(* IEC 61131-3 sources: botanik2/src/libbotanik/plc/functions, 5 files *)

(* ---- health.st ---- *)
(* What a program says about its own answer
   ------------------------------------------------------------------------ *)

(* The codes are Plc::Health's, in its order: matiec numbers an enumeration
   0,1,2... in declaration order, and the two sides have to agree because the
   value IS the program's health row. matiec rejects explicit values here, so
   the order is the contract.

   Only a program that OPTS IN (`health` in programs.csv) has a row to write,
   and one that opts in owes a write to it on every path - which the generator
   checks off matiec's own write list, the same way it checks a quality.

   Every output is written on every scan, so this is never about whether a row
   moved. It is what the number MEANS. *)

TYPE
  HEALTH : (HEALTHY, DEGRADED, FAULTED);
END_TYPE

FUNCTION WORST_HEALTH : HEALTH
(* How a program that leans on another's answer inherits it: the weaker of the
   two. Spelled as comparisons rather than as a maximum, because the ordering
   of an enumerated type is not something to lean on. *)
VAR_INPUT
  A : HEALTH;
  B : HEALTH;
END_VAR
  IF A = FAULTED OR B = FAULTED THEN WORST_HEALTH := FAULTED;
  ELSIF A = DEGRADED OR B = DEGRADED THEN WORST_HEALTH := DEGRADED;
  ELSE WORST_HEALTH := HEALTHY; END_IF;
END_FUNCTION

FUNCTION VERDICT : HEALTH
(* The common shape, said once: whether the law could answer at all, and
   whether it trusted what it answered on.

   ANSWERED is asked first and separately because the two are not degrees of
   one thing: a law with no evidence at all writes its safe state, which is a
   different fact from a law that chose a fallback and stands behind it. *)
VAR_INPUT
  ANSWERED : BOOL;
  TRUSTED  : BOOL;
END_VAR
  IF NOT ANSWERED THEN VERDICT := FAULTED;
  ELSIF NOT TRUSTED THEN VERDICT := DEGRADED;
  ELSE VERDICT := HEALTHY; END_IF;
END_FUNCTION

(* ---- quality.st ---- *)
(* What a reading is worth, and the two ways a law asks
   ------------------------------------------------------------------------ *)

(* The codes are Vars::Quality's, in its order: matiec numbers an enumeration
   0,1,2... in declaration order, and the two sides have to agree because the
   value IS the companion row's. matiec rejects explicit values here, so the
   order is the contract.

   Three, and each is a DECISION a reader makes differently: nothing behind the
   row, something measured, or a number the law stands behind though nothing
   measured it. The reasons a reading went bad - stale, out of band, refused -
   are diagnoses rather than decisions, and each has a home of its own: the
   stamp's age, the band beside the value, and one log line from the master. *)

TYPE
  QUALITY : (Q_NONE, Q_GOOD, Q_HELD);
END_TYPE

FUNCTION GOOD : BOOL
(* Whether something MEASURED it. What a law gating on seeing the plant asks. *)
VAR_INPUT
  Q : QUALITY;
END_VAR
  GOOD := Q = Q_GOOD;
END_FUNCTION

FUNCTION USABLE : BOOL
(* Whether there is a NUMBER behind it worth computing on. Wider than GOOD by
   exactly Q_HELD, which is a law's own fallback. *)
VAR_INPUT
  Q : QUALITY;
END_VAR
  USABLE := Q <> Q_NONE;
END_FUNCTION

FUNCTION WORST_OF : QUALITY
(* How a derived row inherits its inputs': the weaker of the two. Spelled as
   comparisons rather than as a minimum, because the ordering of an enumerated
   type is not something to lean on. *)
VAR_INPUT
  A : QUALITY;
  B : QUALITY;
END_VAR
  IF A = Q_NONE OR B = Q_NONE THEN WORST_OF := Q_NONE;
  ELSIF A = Q_HELD OR B = Q_HELD THEN WORST_OF := Q_HELD;
  ELSE WORST_OF := Q_GOOD; END_IF;
END_FUNCTION

FUNCTION QUAL : QUALITY
(* The quality of a row a law publishes with no input verdict to inherit:
   measured this beat, HOLDING something it measured once, or nothing it has
   ever seen.

   SEEDED is asked separately and always, because the middle case is the one
   that gets skipped: a block whose output holds its last reading and reports
   only OK publishes Q_NONE for a row that has real evidence in it, and
   Ref::get() then hands every reader the declared value instead. Pass FALSE
   where the law genuinely holds nothing - a verdict recomputed each scan - and
   let that be a claim somebody made rather than a default. *)
VAR_INPUT
  OK     : BOOL;
  SEEDED : BOOL;
END_VAR
  IF OK THEN QUAL := Q_GOOD;
  ELSIF SEEDED THEN QUAL := Q_HELD;
  ELSE QUAL := Q_NONE; END_IF;
END_FUNCTION

(* ---- math.st ---- *)
(* The demand ladders, and the votes a redundant chain reduces with
   ------------------------------------------------------------------------ *)

(* Written once so three subsystems cannot disagree about what "half demand"
   means. Stateless, so FUNCTIONs rather than blocks. *)

FUNCTION LADDER : REAL
(* V mapped onto 0..1 across [LO, HI] and clamped. A degenerate or inverted
   span reads as fully on at or above HI, so a mis-set pair fails toward
   ACTING rather than toward doing nothing. *)
VAR_INPUT
  V  : REAL;
  LO : REAL;
  HI : REAL;
END_VAR
  IF HI <= LO THEN
    IF V >= HI THEN LADDER := 1.0; ELSE LADDER := 0.0; END_IF;
  ELSE
    LADDER := LIMIT(0.0, (V - LO) / (HI - LO), 1.0);
  END_IF;
END_FUNCTION

FUNCTION SIGNED_LADDER : REAL
(* The same either side of zero, with a dead band between. Reads 0 inside
   [NEG_START, POS_START], falls to -1 by NEG_FULL and rises to +1 by
   POS_FULL. One signed number, negative meaning the opposite process. *)
VAR_INPUT
  V         : REAL;
  NEG_FULL  : REAL;
  NEG_START : REAL;
  POS_START : REAL;
  POS_FULL  : REAL;
END_VAR
  IF V >= POS_START THEN
    SIGNED_LADDER := LADDER(V := V, LO := POS_START, HI := POS_FULL);
  ELSIF V <= NEG_START THEN
    SIGNED_LADDER := -LADDER(V := -V, LO := -NEG_START, HI := -NEG_FULL);
  ELSE
    SIGNED_LADDER := 0.0;
  END_IF;
END_FUNCTION

FUNCTION MEDIAN3 : REAL
(* The middle of three readings, so one stuck high or stuck low can never be
   the one retained. Both extremes are discarded, not averaged in. *)
VAR_INPUT
  A : REAL;
  B : REAL;
  C : REAL;
END_VAR
  IF   (A <= B AND B <= C) OR (C <= B AND B <= A) THEN MEDIAN3 := B;
  ELSIF (B <= A AND A <= C) OR (C <= A AND A <= B) THEN MEDIAN3 := A;
  ELSE MEDIAN3 := C;
  END_IF;
END_FUNCTION

FUNCTION AVG2 : REAL
(* The mean of two readings: what is left when there is no middle to keep. *)
VAR_INPUT
  A : REAL;
  B : REAL;
END_VAR
  AVG2 := 0.5 * (A + B);
END_FUNCTION

(* ---- psychro.st ---- *)
(* Psychrometrics: dew points, and the margin to them
   ------------------------------------------------------------------------ *)

(* DEW POINTS, not humidities: air at 90% and 5 degC is drier than air at 60%
   and 25, and swapping one for the other is what ventilating does. *)

FUNCTION DEW_POINT : REAL
(* The temperature at which this air saturates and its vapour begins
   condensing onto whatever it touches. Magnus, valid -40..+50 degC.
   RH is a FRACTION, 0..1, never a percentage. *)
VAR_INPUT
  T_DEGC : REAL;
  RH     : REAL;
END_VAR
VAR
  gamma : REAL;
END_VAR
  (* The floor keeps the logarithm defined: bone-dry air is not a reason to
     return minus infinity to a control law. *)
  gamma := LN(LIMIT(0.05, RH, 1.0)) + (17.62 * T_DEGC) / (243.12 + T_DEGC);
  DEW_POINT := (243.12 * gamma) / (17.62 - gamma);
END_FUNCTION

FUNCTION DEW_POINT_MARGIN : REAL
(* How far the air is from condensing, in degC. LARGER is drier. What the rot
   and condensation laws are set in, because it is the margin that decides
   whether water lands on a plant at the temperature it is actually at. *)
VAR_INPUT
  T_DEGC : REAL;
  RH     : REAL;
END_VAR
  DEW_POINT_MARGIN := T_DEGC - DEW_POINT(T_DEGC := T_DEGC, RH := RH);
END_FUNCTION

FUNCTION SAT_VAPOUR_PRESSURE : REAL
(* The most water this air could hold, in kPa. Tetens, whose coefficients are
   NOT Magnus's above: mixing the two sets shifts the answer. *)
VAR_INPUT
  T_DEGC : REAL;
END_VAR
  SAT_VAPOUR_PRESSURE := 0.6108 * EXP((17.27 * T_DEGC) / (T_DEGC + 237.3));
END_FUNCTION

(* ---- time.st ---- *)
(* Seconds as milliseconds, the one place the factor is written
   ------------------------------------------------------------------------ *)

(* A parameter an operator sets is in SECONDS; every timer input is in
   milliseconds. This is that seam, named once, so no law spells the factor
   out and none of them can spell it differently. *)

FUNCTION SEC_MS : UDINT
VAR_INPUT
  S : UINT;
END_VAR
  SEC_MS := UINT_TO_UDINT(S) * 1000;
END_FUNCTION
